(*
SPDX-FileCopyrightText: c 2026 Oleksandr Tiutyk <trofimich@gmail.com>
SPDX-License-Identifier: MIT
License: https://opensource.org/license/mit
*)

(*!
<summary>Checks ANY lookup of present and absent values without changing the queue.</summary>
<description>
Owns an inline queue and its copied entry payloads. Run from one task at a stable address.
Teardown clears surviving entries before publication, including after an aborted case.
</description>
*)

{attribute 'no_assign'}
{attribute 'no_explicit_call' := 'do not call this function block directly'}
FUNCTION_BLOCK StaticQueueContainsTest EXTENDS TOF_Testing.SingleCycleTest
VAR_STAT
	{attribute 'hide'}
	_ClassName : STRING := __POUNAME();
END_VAR
VAR
	_Queue : TOF_Collections.Queue<3>(valueValidator := 0);
END_VAR

(*!
<summary>Checks ANY lookup of present and absent values without changing the queue.</summary>
*)
METHOD PROTECTED ExecuteTest
VAR
	values : ARRAY [1..4] OF INT := [11, 22, 33, 44];
END_VAR
Assert.ThatBool(
	actual := _Queue.Contains(value := values[1]),
	message := "An empty queue must report absence"
).IsFalse();

_Queue
	.EnqueueCopy(value := values[1])
	.EnqueueCopy(value := values[2])
	.EnqueueCopy(value := values[3]);

Assert.ThatBool(
	actual := _Queue.Contains(value := values[1]),
	message := "Contains must find the head"
).IsTrue();

Assert.ThatBool(
	actual := _Queue.Contains(value := values[3]),
	message := "Contains must find the tail"
).IsTrue();

Assert.ThatBool(
	actual := _Queue.Contains(value := values[4]),
	message := "Contains must report a missing value"
).IsFalse();

Assert.ThatDInt(
	actual := _Queue.Length,
	message := "Lookup must preserve all three entries"
).ToBe(expected := DINT#3);

Assert.ThatInt(
	actual := _Queue.Peek().AsInt(),
	message := "Lookup must preserve the head"
).ToBe(expected := values[1]);
END_METHOD

(*!
<summary>Restores the fixture before the runner publishes the result.</summary>
<description>
Also runs after an unexpected exception interrupts the case.
</description>
*)
METHOD PROTECTED AfterTest
_Queue.Clear();
END_METHOD

//! <summary>Borrows the concrete class name. Callers must not modify it.</summary>
{attribute 'monitoring' := 'call'}
PROPERTY ClassName : REFERENCE TO STRING
GET
ClassName REF= _ClassName;
END_GET
END_PROPERTY

//! <summary>Borrows the compiler-initialized namespace name. Callers must not modify it.</summary>
{attribute 'monitoring' := 'call'}
PROPERTY NamespaceName : REFERENCE TO STRING
GET
NamespaceName REF= CurrentNamespace.Name;
END_GET
END_PROPERTY

//! <summary>Reports the concrete instance size in bytes.</summary>
{attribute 'monitoring' := 'call'}
PROPERTY SelfSize : ULINT
GET
SelfSize := XSIZEOF(THIS^);
END_GET
END_PROPERTY

END_FUNCTION_BLOCK

(* stored: Version 1.1.0.1
   POU StaticQueueContainsTest: Id {10eb6bdf-ff45-45cb-814e-bc35f9f88036}, SpecialFunc None
   Method ExecuteTest: Id {6ca08d75-b40f-41ee-a222-a410ec11da41}
   Method AfterTest: Id {882b8915-1cd2-4693-9f98-ac13e60f97cf}
   Property ClassName: Id {94ca1d4e-ce19-437e-b189-2cfedc11d638}
   Get Get: Id {536cc435-ae5e-414e-9896-a528d704588e}
   Property NamespaceName: Id {577a2ee3-20ad-4e67-8c4e-52618332b258}
   Get Get: Id {4344842d-3c34-470a-95bf-73c6eacad22d}
   Property SelfSize: Id {da181fa0-28d0-4761-9633-70760fa6c31f}
   Get Get: Id {346f628c-7619-40e7-9e71-13d09df74cbe} *)
